// TIA Portal V21 export
// export: Created 2026-11-10T07:35:26.7443645Z, ExportSetting WithDefaults, DisplayName Totally Integrated Automation Portal, DisplayVersion V21 Update 3, DisplayName STEP 7 Professional, DisplayVersion V21 Update 3, DisplayName STEP 7 Safety, DisplayVersion V21, DisplayName Tech WebApplication, DisplayVersion V21, DisplayName WinCC Basic/Comfort/Advanced, DisplayVersion V21 Update 3, DisplayName WinCC Unified, DisplayVersion V21 Update 3
FUNCTION_BLOCK "FB_Lad_ou015"   // FB81, LAD
{ S7_Optimized_Access := 'TRUE' }
VERSION : 0.1
// stored: AutoNumber true, IsIECCheckEnabled false, IsRetainMemResEnabled false, MemoryReserve 100, SetENOAutomatically false, UDAEnableTagReadback false
   VAR_INPUT
      v_en_r : Bool;
      v_id : CONN_OUC;
      v_len : UInt;
      v_adhoc : Bool;
   END_VAR
   VAR_OUTPUT
      v_ndr : Bool;
      v_busy : Bool;
      v_error : Bool;
      v_status : Word;
      v_rcvd_len : UInt;
   END_VAR
   VAR_IN_OUT
      v_data : Array[0..99] of Byte;
   END_VAR
   VAR
      inst { S7_SetPoint := 'True'} : TRCV;
   END_VAR
BEGIN

REGION Network 1: TRCV - Receive data via communication connection
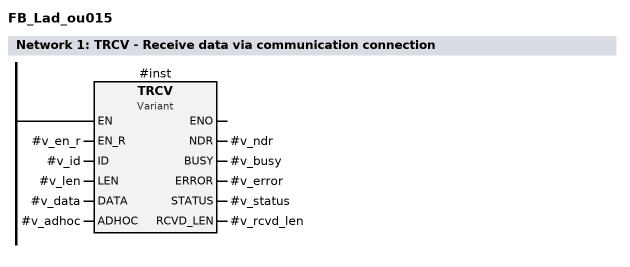
   RUNG wire#powerrail
      { S7_Templates := "[card := 1, ptr_type := Variant, value_type := UDInt, id_type := CONN_OUC]" } #inst.TRCV(EN_R := #v_en_r, ID := #v_id, LEN := #v_len, DATA := #v_data, NDR => #v_ndr, BUSY => #v_busy, ERROR => #v_error, STATUS => #v_status, RCVD_LEN => #v_rcvd_len, ADHOC := #v_adhoc)
   END_RUNG
   // the same network as SCL:
   #inst(EN_R := #v_en_r,   // TRCV
         ID := #v_id,
         LEN := #v_len,
         DATA := #v_data,
         ADHOC := #v_adhoc,
         NDR => #v_ndr,
         BUSY => #v_busy,
         ERROR => #v_error,
         STATUS => #v_status,
         RCVD_LEN => #v_rcvd_len);
END_REGION
END_FUNCTION_BLOCK
